FUNCTION_BLOCK FB_3002_ModbusTcpClient
(* ==============================================================================
 * FB_3002_ModbusTcpClient - 上下游 Modbus TCP 客户端数据映射层
 * 项目: DJ-2026-009 汇川换型改造
 * 依据: BC-DJ-2026-009-004, 通讯契约 V0.3 (030_DJ-2026-009_通讯契约_INT.md) 2.0~2.2
 * 实施卡: CARD-DJ-2026-009-001
 *
 * 职责:
 *   本机做 Modbus TCP 客户端. 报文收发由 InoProShop 的 Modbus TCP 主站通道完成,
 *   通道把对方保持寄存器映射到 4 个寄存器镜像数组 (下标 = 协议地址, 从 0 起).
 *   本块只做两件事:
 *     1. 把读回的镜像解包到 ST_UpstreamDocking / ST_DownstreamDocking (对方 -> 本机);
 *        把本机信号封包到写镜像 (本机 -> 对方).
 *     2. 根据通道链路状态给出通讯状态位和错误码.
 *   链路断开时读侧变量保持最后值不刷新, 心跳因此停止翻转,
 *   由 FB_3001 现有的 12s 心跳超时照常报通讯故障. 本块不直接改握手状态.
 *
 * STRING 按字符取下标: 下标从 1 起 (第 1 个字符是 s[1])。这是 siemens-lsp 插件 (S7 语义) 的要求;
 *   移植到汇川 InoProShop / CODESYS 等平台须按平台适配 (这类平台字符下标可能从 0 起)。
 *   适配点: 本文件里所有 s_sIdBuf[...] 的下标 (组件 ID 解包 3 处、封包 2 处), 数组下标不受影响。
 *
 * 寄存器地址取自契约 V0.3 我方提议版, 未经对方签字, 见下方 VAR CONSTANT.
 * ============================================================================== *)
VAR_INPUT
    i_bEnable           : BOOL;         // 功能块总使能
    i_bUpLinkOK         : BOOL;         // 上游 Modbus TCP 通道链路正常 (来自主站通道诊断)
    i_bDownLinkOK       : BOOL;         // 下游 Modbus TCP 通道链路正常 (来自主站通道诊断)
END_VAR

VAR_OUTPUT
    q_bComOK            : BOOL;         // 上下游通道链路均正常
    q_wErrorCode        : WORD;         // 通讯层故障诊断字 (bit0 上游链路断, bit1 下游链路断)
END_VAR

VAR_IN_OUT
    io_stExternal       : ST_ExternalDevice;        // STD-820 通用外部对接数据总线
    io_arrUpRead        : ARRAY[0..31] OF WORD;     // 上游寄存器读镜像 (下标 = 协议地址)
    io_arrUpWrite       : ARRAY[0..31] OF WORD;     // 上游寄存器写镜像 (下标 = 协议地址)
    io_arrDownRead      : ARRAY[0..31] OF WORD;     // 下游寄存器读镜像 (下标 = 协议地址)
    io_arrDownWrite     : ARRAY[0..31] OF WORD;     // 下游寄存器写镜像 (下标 = 协议地址)
END_VAR

VAR
    s_wStatusIn         : WORD;         // 解包用: 对方状态字
    s_wStatusOut        : WORD;         // 封包用: 本机状态字
    s_iReg              : INT;          // 组件 ID 寄存器循环下标 (0~15)
    s_iChar             : INT;          // 组件 ID 字符下标 (0~31)
    s_bIdEnd            : BOOL;         // 解包组件 ID 时已遇到结束符 0
    s_byHi              : BYTE;         // 寄存器高字节 (前一个字符)
    s_byLo              : BYTE;         // 寄存器低字节 (后一个字符)
    s_sIdBuf            : STRING[32];   // 组件 ID 解包缓冲
    s_wErrorCode        : WORD;         // 通讯层故障诊断字 (内部累加, 块内判断用, 块末尾赋给输出 q_wErrorCode)
END_VAR

VAR CONSTANT
    // --- 寄存器地址 (契约 V0.3 2.0, 我方提议, 待对方签字) ---
    REG_STATUS_IN       : INT := 0;     // 对方 -> 本机 状态字
    REG_STATUS_OUT      : INT := 1;     // 本机 -> 对方 状态字
    REG_ID_START        : INT := 2;     // 组件 ID 起始地址 (2~17 共 16 个寄存器)
    ID_REG_COUNT        : INT := 16;    // 组件 ID 寄存器个数 (32 字符 / 2)
    REG_IMAGE_LAST      : INT := 31;    // 镜像数组最后一个下标 (18~31 预留)

    // --- 状态字位掩码 (bit0 为最低位) ---
    MASK_B0             : WORD := 16#0001;
    MASK_B1             : WORD := 16#0002;
    MASK_B2             : WORD := 16#0004;
    MASK_B3             : WORD := 16#0008;
    MASK_B15            : WORD := 16#8000;  // 心跳位

    // --- 错误码 ---
    ERR_NONE            : WORD := 16#0000;
    ERR_UP_LINK         : WORD := 16#0001;  // 上游通道链路断开
    ERR_DOWN_LINK       : WORD := 16#0002;  // 下游通道链路断开
END_VAR

BEGIN
    IF NOT i_bEnable THEN
        // 未使能: 本机发给对方的状态字和组件 ID 全部清零 (对方看到的允许/请求信号均为 0)
        FOR s_iReg := 0 TO REG_IMAGE_LAST DO
            io_arrUpWrite[s_iReg] := 16#0000;
            io_arrDownWrite[s_iReg] := 16#0000;
        END_FOR;
        q_bComOK := FALSE;
        q_wErrorCode := ERR_NONE;
        RETURN;
    END_IF;

    (* 1. 链路状态与错误码 *)
    s_wErrorCode := ERR_NONE;
    IF NOT i_bUpLinkOK THEN
        s_wErrorCode := s_wErrorCode OR ERR_UP_LINK;
    END_IF;
    IF NOT i_bDownLinkOK THEN
        s_wErrorCode := s_wErrorCode OR ERR_DOWN_LINK;
    END_IF;
    // 输出只在此处赋值, 块内不再读取输出参数 (TIA 对读输出参数报警)。
    q_wErrorCode := s_wErrorCode;
    q_bComOK := (s_wErrorCode = ERR_NONE);

    (* 2. 上游读解包 (链路断开时保持最后值, 由 FB_3001 心跳超时判故障) *)
    IF i_bUpLinkOK THEN
        s_wStatusIn := io_arrUpRead[REG_STATUS_IN];
        io_stExternal.stUpstream.bUpstream_LineReady := (s_wStatusIn AND MASK_B0) <> 16#0000;
        io_stExternal.stUpstream.bUpstream_SendModuleId := (s_wStatusIn AND MASK_B1) <> 16#0000;
        io_stExternal.stUpstream.bUpstream_InfeedReq := (s_wStatusIn AND MASK_B2) <> 16#0000;
        io_stExternal.stUpstream.bUpstream_InfeedArrivedAck := (s_wStatusIn AND MASK_B3) <> 16#0000;
        io_stExternal.stUpstream.bUpstream_HeartbeatFromUp := (s_wStatusIn AND MASK_B15) <> 16#0000;

        // 组件 ID: 每个寄存器 2 个字符, 高字节在前; 遇到 0 即结束, 内容原样保留
        s_sIdBuf := '';
        s_bIdEnd := FALSE;
        s_iChar := 0;
        FOR s_iReg := 0 TO ID_REG_COUNT - 1 DO
            s_byHi := WORD_TO_BYTE(SHR(io_arrUpRead[REG_ID_START + s_iReg], 8));
            s_byLo := WORD_TO_BYTE(io_arrUpRead[REG_ID_START + s_iReg] AND 16#00FF);
            IF NOT s_bIdEnd THEN
                IF s_byHi = 16#00 THEN
                    s_bIdEnd := TRUE;
                ELSE
                    s_sIdBuf[s_iChar + 1] := s_byHi;  // STRING 下标从 1 起，为 siemens-lsp 插件（S7 语义）要求；移植到汇川 InoProShop / CODESYS 等平台须按平台适配
                    s_iChar := s_iChar + 1;
                END_IF;
            END_IF;
            IF NOT s_bIdEnd THEN
                IF s_byLo = 16#00 THEN
                    s_bIdEnd := TRUE;
                ELSE
                    s_sIdBuf[s_iChar + 1] := s_byLo;  // STRING 下标从 1 起，为 siemens-lsp 插件（S7 语义）要求；移植到汇川 InoProShop / CODESYS 等平台须按平台适配
                    s_iChar := s_iChar + 1;
                END_IF;
            END_IF;
        END_FOR;
        // 按下标逐字符写入不会更新字符串当前长度 (S7 语义): 把长度截到实际字符数 (结束符由字符串自带, 不再手写, 32 个字符满时也不越界)
        s_sIdBuf := LEFT(s_sIdBuf, s_iChar);
        io_stExternal.stUpstream.sRcvModuleID := s_sIdBuf;
    END_IF;

    (* 3. 下游读解包 (链路断开时保持最后值) *)
    IF i_bDownLinkOK THEN
        s_wStatusIn := io_arrDownRead[REG_STATUS_IN];
        io_stExternal.stDownstream.bDownstream_LineReady := (s_wStatusIn AND MASK_B0) <> 16#0000;
        io_stExternal.stDownstream.bDownstream_RcvModuleIdAck := (s_wStatusIn AND MASK_B1) <> 16#0000;
        io_stExternal.stDownstream.bDownstream_AllowOutfeed := (s_wStatusIn AND MASK_B2) <> 16#0000;
        io_stExternal.stDownstream.bDownstream_OutfeedArrived := (s_wStatusIn AND MASK_B3) <> 16#0000;
        io_stExternal.stDownstream.bDownstream_HeartbeatFromDown := (s_wStatusIn AND MASK_B15) <> 16#0000;
    END_IF;

    (* 4. 上游写封包: 本机 -> 上游 状态字 (地址 1), 未用位填 0 *)
    s_wStatusOut := 16#0000;
    IF io_stExternal.stUpstream.bMachine_ReadyIn THEN
        s_wStatusOut := s_wStatusOut OR MASK_B0;
    END_IF;
    IF io_stExternal.stUpstream.bMachine_RcvModuleIdAck THEN
        s_wStatusOut := s_wStatusOut OR MASK_B1;
    END_IF;
    IF io_stExternal.stUpstream.bMachine_AllowInfeed THEN
        s_wStatusOut := s_wStatusOut OR MASK_B2;
    END_IF;
    IF io_stExternal.stUpstream.bMachine_InfeedArrived THEN
        s_wStatusOut := s_wStatusOut OR MASK_B3;
    END_IF;
    IF io_stExternal.stUpstream.bMachine_HeartbeatToUp THEN
        s_wStatusOut := s_wStatusOut OR MASK_B15;
    END_IF;
    io_arrUpWrite[REG_STATUS_OUT] := s_wStatusOut;

    (* 5. 下游写封包: 本机 -> 下游 状态字 (地址 1) 与组件 ID (地址 2~17) *)
    s_wStatusOut := 16#0000;
    IF io_stExternal.stDownstream.bMachine_ReadyOut THEN
        s_wStatusOut := s_wStatusOut OR MASK_B0;
    END_IF;
    IF io_stExternal.stDownstream.bMachine_SendModuleId THEN
        s_wStatusOut := s_wStatusOut OR MASK_B1;
    END_IF;
    IF io_stExternal.stDownstream.bMachine_OutfeedReq THEN
        s_wStatusOut := s_wStatusOut OR MASK_B2;
    END_IF;
    IF io_stExternal.stDownstream.bMachine_OutfeedArrivedAck THEN
        s_wStatusOut := s_wStatusOut OR MASK_B3;
    END_IF;
    IF io_stExternal.stDownstream.bMachine_HeartbeatToDown THEN
        s_wStatusOut := s_wStatusOut OR MASK_B15;
    END_IF;
    io_arrDownWrite[REG_STATUS_OUT] := s_wStatusOut;

    // 组件 ID 原样封包: 第 2n 个字符放高字节, 第 2n+1 个放低字节, 不足 32 个字符补 0
    s_sIdBuf := io_stExternal.stDownstream.sSendModuleID;
    s_iChar := LEN(s_sIdBuf);
    FOR s_iReg := 0 TO ID_REG_COUNT - 1 DO
        s_byHi := 16#00;
        s_byLo := 16#00;
        IF (2 * s_iReg) < s_iChar THEN
            s_byHi := s_sIdBuf[2 * s_iReg + 1];  // STRING 下标从 1 起，为 siemens-lsp 插件（S7 语义）要求；移植到汇川 InoProShop / CODESYS 等平台须按平台适配
        END_IF;
        IF (2 * s_iReg + 1) < s_iChar THEN
            s_byLo := s_sIdBuf[2 * s_iReg + 2];  // STRING 下标从 1 起，为 siemens-lsp 插件（S7 语义）要求；移植到汇川 InoProShop / CODESYS 等平台须按平台适配
        END_IF;
        io_arrDownWrite[REG_ID_START + s_iReg] := SHL(BYTE_TO_WORD(s_byHi), 8) OR BYTE_TO_WORD(s_byLo);
    END_FOR;

END_FUNCTION_BLOCK
